(* IEC 61131-3 sources: SRCI_CLIENT_PLC/RobotLibrary/Library/POUs/Read/MC_ReadMessages/Structures, 4 files *)

(* ---- ReadMessagesOutCmd.st ---- *)
{attribute 'pack_mode' := '1'}
// -------------------------------------------------------------------------
//  SRCI Robot Library
// -------------------------------------------------------------------------
//
//  Object:      ReadMessagesOutCmd
//  Author:      Thorsten Brach
//  Date:        2024-08-09
//
//  Description:
//
//
//  Copyright:
//    (C) 2024 Thorsten Brach. All rights reserved
//             Licensed under the MIT License.
//
//  Disclaimer:
//    This project is provided without any guarantee and can be used for
//    private and commercial purposes. Any use is at the user’s
//    own risk and responsibility.
//
// -------------------------------------------------------------------------
TYPE ReadMessagesOutCmd :
STRUCT
  /// ID for function specific acknowledgement mechanism
  MsgId                  : USINT;
  /// Number of pending errors on RC
  NumberOfActiveErrors   : USINT;
  /// Number if pending warnings in RC
  NumberOfActiveWarnings : USINT;
  /// Timestamp
  Timestamp              : IEC_TIMESTAMP;
  /// Message Type
  MsgType                : MessageType;
  /// Severity of returned message according to .Table 5-49.
  Severity               : Severity;
  /// ErrorCode
  ErrorCode              : DWORD;
  /// Test
  Text                   : STRING(255);
END_STRUCT
END_TYPE

(* ---- ReadMessagesParCmd.st ---- *)
{attribute 'pack_mode' := '1'}
// -------------------------------------------------------------------------
//  SRCI Robot Library
// -------------------------------------------------------------------------
//
//  Object:      ReadMessagesParCmd
//  Author:      Thorsten Brach
//  Date:        2024-08-09
//
//  Description:
//
//
//  Copyright:
//    (C) 2024 Thorsten Brach. All rights reserved
//             Licensed under the MIT License.
//
//  Disclaimer:
//    This project is provided without any guarantee and can be used for
//    private and commercial purposes. Any use is at the user’s
//    own risk and responsibility.
//
// -------------------------------------------------------------------------
TYPE ReadMessagesParCmd :
STRUCT
  /// ID for function specific acknowledgement mechanism
  MsgID        : USINT;
  /// Defines up to which level of severity messages will be transmitted to the PLC’s message buffer
  MessageLevel : MessageLevel;
END_STRUCT
END_TYPE

(* ---- ReadMessagesRecvData.st ---- *)
{attribute 'pack_mode' := '1'}
// -------------------------------------------------------------------------
//  SRCI Robot Library
// -------------------------------------------------------------------------
//
//  Object:      ReadMessagesRecvData
//  Author:      Thorsten Brach
//  Date:        2024-08-09
//
//  Description:
//
//
//  Copyright:
//    (C) 2024 Thorsten Brach. All rights reserved
//             Licensed under the MIT License.
//
//  Disclaimer:
//    This project is provided without any guarantee and can be used for
//    private and commercial purposes. Any use is at the user’s
//    own risk and responsibility.
//
// -------------------------------------------------------------------------
TYPE ReadMessagesRecvData EXTENDS RspHeader :
STRUCT
  /// Set TRUE to read messages from RC.
  Enabled                : BOOL;
  /// ID for function specific acknowledgement mechanism
  MsgId                  : USINT;
  /// Number of pending errors on RC
  NumberOfActiveErrors   : USINT;
  /// Number if pending warnings in RC
  NumberOfActiveWarnings : USINT;
  /// Timestamp
  Timestamp              : IEC_TIMESTAMP;
  /// Message Type
  MsgType                : USINT;
  /// Severity of returned message according to .Table 5-49.
  Severity               : SINT;
  /// ErrorCode
  ErrorCode              : DWORD;
  /// Test
  Text                   : STRING(255);
END_STRUCT
END_TYPE

(* ---- ReadMessagesSendData.st ---- *)
{attribute 'pack_mode' := '1'}
// -------------------------------------------------------------------------
//  SRCI Robot Library
// -------------------------------------------------------------------------
//
//  Object:      ReadMessagesSendData
//  Author:      Thorsten Brach
//  Date:        2024-08-09
//
//  Description:
//
//
//  Copyright:
//    (C) 2024 Thorsten Brach. All rights reserved
//             Licensed under the MIT License.
//
//  Disclaimer:
//    This project is provided without any guarantee and can be used for
//    private and commercial purposes. Any use is at the user’s
//    own risk and responsibility.
//
// -------------------------------------------------------------------------
TYPE ReadMessagesSendData EXTENDS CmdHeader:
STRUCT
  /// ID for function specific acknowledgement mechanism
  MsgID        : USINT;
  /// TRUE when function is returning messages from RC
  Enable       : BOOL;
  /// Defines up to which level of severity messages will be transmitted to the PLC’s message buffer
  MessageLevel : USINT;
END_STRUCT
END_TYPE
